       ELSIF (#tempEnable = FALSE) AND (#statEnableOld = TRUE) THEN // Disable FB 
           #statFBState := #FB_STATE_DISABLING;
       ELSIF (#statStatus = #STATUS_FIRST_CALL) THEN // Set status identifier of subsequent call
           #statStatus := #STATUS_SUBSEQUENT_CALL;
       END_IF;

       // Edge detection 'enable' input
       #statEnableOld := #tempEnable;
   END_REGION ENABLING/DISABLING

   IF (#statStatus = #STATUS_NO_CALL) THEN // Nothing to do -> End here to reduce "system load"
       RETURN;
   END_IF;

   REGION STATE_MACHINE_FUNCTION_BLOCK_TCP
       CASE #statFBState OF // State machine of FB
           #FB_STATE_NO_PROCESSING: // No processing active (Note: this state must always be present and left empty)
               ;

           #FB_STATE_VALIDATE_INPUT: // Enabling active
               REGION EVALUATE CONNECTION PARAMETERS
                   // Determine if host is domain name or IP address
                   #statConnParam.isQDN := NOT "IsIPAddress"(address := #connParam.broker, ipAddress => #statConnParam.paramIP.ConnPara.RemoteAddress);

                   IF #statConnParam.isQDN THEN // Broker address is a hostname
                       IF #connParam.broker[LEN(#connParam.broker)] = '.' THEN
                           #statConnParam.paramQDN.ConnPara.RemoteQDN := #connParam.broker;
                       ELSE
                           #statConnParam.paramQDN.ConnPara.RemoteQDN := CONCAT(IN1 := #connParam.broker, IN2 := '.');
                       END_IF;

                       #statConnParam.paramQDN.ConnPara.InterfaceId := #connParam.hwId;
                       #statConnParam.paramQDN.ConnPara.ID := #connParam.connId;
                       #statConnParam.paramQDN.ConnPara.ActiveEstablished := TRUE;
                       #statConnParam.paramQDN.ConnPara.RemotePort := #connParam."port";
                   ELSE // Broker address is an IP address
                       #statConnParam.paramIP.ConnPara.InterfaceId := #connParam.hwId;
                       #statConnParam.paramIP.ConnPara.ID := #statConnParam.paramQDN.ConnPara.ID := #connParam.connId;
                       #statConnParam.paramIP.ConnPara.ActiveEstablished := TRUE;
                       #statConnParam.paramIP.ConnPara.RemotePort := #connParam."port";
                   END_IF;

                   IF #connParam.tls.enableTls THEN
                       IF #statConnParam.isQDN THEN
                           #statConnParam.paramQDN.ActivateSecureConn := TRUE;
                           #statConnParam.paramQDN.ExtTLSCapabilities.%X0 := #connParam.tls.validateServerIdentity;
                           #statConnParam.paramQDN.TLSServerCertRef := #connParam.tls.brokerCert;
                           #statConnParam.paramQDN.TLSClientCertRef := #connParam.tls.clientCert;
                       ELSE
                           #statConnParam.paramIP.ActivateSecureConn := TRUE;
                           #statConnParam.paramIP.ExtTLSCapabilities.%X0 := #connParam.tls.validateServerIdentity;
                           #statConnParam.paramIP.TLSServerCertRef := #connParam.tls.brokerCert;
                           #statConnParam.paramIP.TLSClientCertRef := #connParam.tls.clientCert;
                       END_IF;
                   ELSE
                       IF #statConnParam.isQDN THEN
                           #statConnParam.paramQDN.ActivateSecureConn := FALSE;
                       ELSE
                           #statConnParam.paramIP.ActivateSecureConn := FALSE;
                       END_IF;
                   END_IF;
               END_REGION EVALUATE CONNECTION PARAMETERS

               REGION FB_VALIDATE_INPUT     
                   // Check Input variables:
                   #tempMaxWillMsgLen := ABS(UPPER_BOUND(ARR := #willMsgPayload, DIM := #ONE_DIMENSION) - LOWER_BOUND(ARR := #willMsgPayload, DIM := #ONE_DIMENSION)) + #ARRAY_LEN_OFFSET_PLUS_1;

                   // Check Client ID len Must be > 0 
                   IF LEN(#clientIdentifier) <= #LEN_NULL THEN
                       #statStatus := #ERR_CLIENT_ID_NULL; // Set correct status that identifies error clearly
                       #statSubfunctionStatus := #ERR_CLIENT_ID_NULL; // Status or return value of called FBs, FCs and system blocks
                       #statFBErrorState := #statFBState; // Set error state number for diagnostic 
                       #statErrorUserCleared := TRUE;

                       // Verify Will next
                   ELSIF #tempMaxWillMsgLen < #willMsgLen THEN
                       #statStatus := #ERR_CNT_EXCEEDS_ARRAY_DIMENSION; // Set correct status that identifies error clearly
                       #statSubfunctionStatus := #ERR_CNT_EXCEEDS_ARRAY_DIMENSION; // Status or return value of called FBs, FCs and system blocks
                       #statFBErrorState := #statFBState; // Set error state number for diagnostic 
                       #statErrorUserCleared := TRUE;

                       // Check Will QoS
                   ELSIF #qos > #MQTT_QOS_2 THEN
                       #statStatus := #ERR_QOS_INVALID; // Set correct status that identifies error clearly
                       #statSubfunctionStatus := #ERR_QOS_INVALID; // Status or return value of called FBs, FCs and system blocks
                       #statFBErrorState := #statFBState; // Set error state number for diagnostic 
                       #statErrorUserCleared := TRUE;

                       // Check KeepAlive
                   ELSIF (#connParam.keepAlive < #THREE_SECONDS) // IF Set to 1 or 2 seconds..
                       AND (#connParam.keepAlive > 0)
                   THEN
                       #statStatus := #ERR_KEEPALIVE_INVALID; // Set correct status that identifies error clearly
                       #statSubfunctionStatus := #ERR_KEEPALIVE_INVALID; // Status or return value of called FBs, FCs and system blocks
                       #statFBErrorState := #statFBState; // Set error state number for diagnostic 
                       #statErrorUserCleared := TRUE;

                   ELSE
                       // Set Params for connection
                       // Set Client Id
                       #statWillQos := #qos;
                       // Set Retain
                       #statWillRetain := #retain;
                       // Will message cnt
                       #statWillMessageCnt := #willMsgLen;

                       // Keepalive
                       IF #connParam.keepAlive = 0 THEN
                           #statMqttKeepAliveUsed := FALSE;
                       ELSE
                           #statMqttKeepAliveUsed := TRUE;
                           // KeepAliveTImer is set to ((Keep Alive converted to seconds) - 2s)
                           #statMqttKeepAliveTime := UINT_TO_TIME((#connParam.keepAlive * #UINT_CONST_1000 - #TWO_SECONDS));
                       END_IF;

                       // rdy to enable TCON
                       #statTsendcEnable := TRUE;
                       #statEnableTimerCommandWatchdog := TRUE;
                       #statFBState := #FB_STATE_TCP_CONNECTING;
                   END_IF;
               END_REGION FB_VALIDATE_INPUT

           #FB_STATE_TCP_CONNECTING: // Wait for TCP to be established
               REGION FB_TCP_CONNECTING
                   // Check process:
                   IF #tempTsendcError = TRUE THEN // when error:
                       #statTsendcEnable := FALSE; // disable TsendC
                       #statEnableTimerCommandWatchdog := FALSE;
                       #statStatus := #ERR_TCON_FAILED; // Set correct status that identifies error clearly
                       #statSubfunctionStatus := #tempTsendcStatus; // Status or return value of called FBs, FCs and system blocks
                       #statFBErrorState := #statFBState; // Set error state number for diagnostic 
                       #statErrorUserCleared := TRUE;

                   ELSIF #tempTsendcStatus = #TSENDC_EST_OK THEN // when successfull:
                       // Communication connection established.
                       #statEnableTimerCommandWatchdog := FALSE;
                       // Monitor Connection
                       #statFBState := #FB_STATE_OPERATING_MONITOR_TCP;
                       // Begin MQTT Connection
                       #statMqttConnectState := #MQTT_CONNECT_STATE_BUILD_PACKET;
                       // set status
                       #statStatus := #STATUS_MQTT_CONNECTING;

                   ELSIF #instTimerCommandWatchdog.Q THEN
                       #statTsendcEnable := FALSE; // disable TsendC
                       #statEnableTimerCommandWatchdog := FALSE;
                       #statStatus := #ERR_TCON_TIMEOUT; // Set correct status that identifies error clearly
                       #statSubfunctionStatus := #ERR_TCON_TIMEOUT; // Status or return value of called FBs, FCs and system blocks
                       #statFBErrorState := #statFBState; // Set error state number for diagnostic 
                       #statErrorUserCleared := TRUE;
                   END_IF;
               END_REGION FB_TCP_CONNECTING

           #FB_STATE_OPERATING_MONITOR_TCP: // Processing active
               REGION FB_OPERATING_MONITOR_TCP
                   // Reset Status on Msg Output - will be set when a new message is completly processed and ready at outputs.
                   #statRcvMsgStatus := #MSG_DECODE_STATUS_NO_NEW_MSG;
                   // Reset TsendC Req from last  cycle Request:
                   #statTsendcReq := FALSE;

                   // Monitor Connection - if disconnect occured:
                   IF ((#tempTsendcStatus > #TSENDC_COM_CLOSED AND #tempTsendcStatus < #TSENDC_EST_OK) // Status connection interupt
                       OR #tempTsendcError = TRUE) // Or error
                       AND #tempTrcvNdr = FALSE // And no new data (to see if broker send information why connection was interrupted)
                   THEN
                       REGION CONNECTION_INTERRUPTED
                           // Status reconnecting
                           // SET MQTT to no operation
                           #statMqttConnectState := #MQTT_CONNECT_STATE_NO_PROCESSING;
                           #statMqttCommandState := #MQTT_COMMAND_STATE_NO_PROCESSING;
                           #statRcvMsgDecodeState := #MSG_DECODE_STATE_NO_PROCESSING;
                           // Reset PUBACK / PUBREC / PUBCOMP
                           #statSendPubAckMsg :=
                           #statSendPubRecMsg :=
                           #statSendPubCompMsg := FALSE;
                           // reset Done bit if still set, regardless of input:
                           #statDone := FALSE;
                           // reset Watchdog
                           #statEnableTimerCommandWatchdog := FALSE;
                           // reset headerEncode
                           #statPacketHeaderEncodeDone := FALSE;
                           // set error  information
                           #statStatus := #ERR_TCP_RECONNECTING; // Set correct status that identifies error clearly
                           #statSubfunctionStatus := #tempTsendcStatus;// Status or return value of called FBs, FCs and system blocks
                           #statFBErrorState := #statFBState; // Set error state number for diagnostic 
                           #statErrorAutoCleared := TRUE;
                           // Wait for reconect - next state
                           #statFBState := #FB_STATE_TCP_RECONNECTING;
                       END_REGION REGION CONNECTION_INTERRUPTED
                   ELSE
                       // Connection is OK
                       // Sending and receiving works 
                       // Check Trcv Buffer for new Data
                       IF #tempTrcvNdr THEN
                           REGION TRCV_NEW_DATA
                               // Evaluate the TrcvBuffer, reset buffer pos to start
                               #tempTrcvBufferPos := 0;

                               // Parse the whole RCV Buffer
                               // While there is data to be processed
                               WHILE ((#tempTrcvBufferPos = UDINT_TO_DINT(#tempTrcvRcvdLen) AND #statRcvMsgDecodeState = #MSG_DECODE_STATE_COMPLETED)
                                   OR #tempTrcvBufferPos < UDINT_TO_DINT(#tempTrcvRcvdLen))
                               DO
                                   // Parse the whole RCV Buffer, check wether header or decoding
                                   IF #statRcvMsgDecodeState = #MSG_DECODE_STATE_NO_PROCESSING THEN
                                       // If no decoding is in progress, look for new message header
                                       #tempRcvMsgTypeCase := #statRcvBuffer[#tempTrcvBufferPos] AND #BIT_MASK_HIGHBITS;
                                   ELSE
                                       // Decode is in progress, go directly to decoding
                                       #tempRcvMsgTypeCase := #MQTT_MSG_DECODING;
                                   END_IF;

                                   CASE #tempRcvMsgTypeCase OF

                                       #MQTT_MSG_TYPE_CONNACK:
                                           REGION RECEIVED_CONACK_PACKET
                                               // Check all CONNACK packet is inside the receive buffer
                                               IF #tempTrcvBufferPos + #BYTE_SIZE_CONNACK <= #MAX_BUFFER_LEN_RCV THEN
                                                   #tempTrcvBufferPos += 1;
                                                   IF #statRcvBuffer[#tempTrcvBufferPos] = #REMAINING_LEN_2 THEN // remainng Length must be 2;
                                                       #tempTrcvBufferPos += 1;
                                                       // byte one is 0000 000X where X is if Session was set, so depending on clean session or not evaluate answer of server
                                                       #statSessionPresent := #statRcvBuffer[#tempTrcvBufferPos] <> #MQTT_NO_SESSION_PRESENT;
                                                       IF (#cleanSession AND NOT #statSessionPresent)
                                                           OR NOT #cleanSession
                                                       THEN
                                                           #tempTrcvBufferPos += 1;
                                                           // VALID Answer, check code
                                                           IF #statRcvBuffer[#tempTrcvBufferPos] = #MQTT_CONNACK_ACCEPTED THEN
                                                               // All good
                                                               #tempTrcvBufferPos += 1;
                                                               #tempMqttConnAckRcvStatus := #RESPONSE_GOOD; // evaluate in MQTT StateMachine Below the response
                                                           ELSE
                                                               // NOT VALID CONNACK from server shows session has a bad return code
                                                               #statStatus := #ERR_MQTT_CONNACK_RETURN_CODE_INVALID; // Set correct status that identifies error clearly
                                                               #statSubfunctionStatus := #statRcvBuffer[#tempTrcvBufferPos]; // Status or return value of called FBs, FCs and system blocks
                                                               #statFBErrorState := #statFBState; // Set error state number for diagnostic 
                                                               #statErrorUserCleared := TRUE;
                                                               // Exit loop
                                                               EXIT;
                                                           END_IF;
                                                       ELSE
                                                           // NOT VALID, CONNACK from server shows session present
                                                           #statStatus := #ERR_MQTT_CONNACK_INVALID_SESSION_FLAG; // Set correct status that identifies error clearly
                                                           #statSubfunctionStatus := #ERR_MQTT_CONNACK_INVALID_SESSION_FLAG; // Status or return value of called FBs, FCs and system blocks
                                                           #statFBErrorState := #statFBState; // Set error state number for diagnostic 
                                                           #statErrorUserCleared := TRUE;
                                                           // Exit loop
                                                           EXIT;
                                                       END_IF;
                                                   ELSE // We got a CONNACK packet, but remaining length was not 2 (Error)
                                                       #statStatus := #ERR_MQTT_REM_LEN_INVALID; // Set correct status that identifies error clearly
                                                       #statSubfunctionStatus := #ERR_MQTT_REM_LEN_INVALID; // Status or return value of called FBs, FCs and system blocks
                                                       #statFBErrorState := #statFBState; // Set error state number for diagnostic 
                                                       #statErrorUserCleared := TRUE;
                                                       // Exit loop
                                                       EXIT;
                                                   END_IF;
                                               ELSE
                                                   // If the CONNACK packed is not fully inside the receive buffer, finish processing
                                                   #statStatus := #ERR_MSG_SKIPPED; // Set correct status that identifies error clearly
                                                   #statSubfunctionStatus := #ERR_MSG_SKIPPED; // Status or return value of called FBs, FCs and system blocks
                                                   #statFBErrorState := #statFBState; // Set error state number for diagnostic 
                                                   #statErrorUserCleared := TRUE;
                                                   // Exit loop
                                                   EXIT;
                                               END_IF;
                                           END_REGION RECEIVED_CONACK_PACKET

                                       #MQTT_MSG_TYPE_PINGRESP:
                                           REGION RECEIVED_PINGRESP_PACKET
                                               // Check all PINGRESP packet is inside the receive buffer
                                               IF #tempTrcvBufferPos + #BYTE_SIZE_PINGRESP <= #MAX_BUFFER_LEN_RCV THEN
                                                   #tempTrcvBufferPos += 1;
                                                   IF #statRcvBuffer[#tempTrcvBufferPos] = #REMAINING_LEN_0 THEN // remainng Length must be 0;
                                                       #tempTrcvBufferPos += 1;
                                                       #tempMqttPingRspRcv := #RESPONSE_GOOD; // evaluate in MQTT StateMachine Below the response
                                                   ELSE // We got a Pingrsp packet, but remaining length was not 0 (Error)
                                                       #statStatus := #ERR_MQTT_REM_LEN_INVALID; // Set correct status that identifies error clearly
                                                       #statSubfunctionStatus := #ERR_MQTT_REM_LEN_INVALID; // Status or return value of called FBs, FCs and system blocks
                                                       #statFBErrorState := #statFBState; // Set error state number for diagnostic 
                                                       #statErrorAutoCleared := TRUE;
                                                       // Exit loop
                                                       EXIT;
                                                   END_IF;
                                               ELSE
                                                   // If the PINGRESP packed is not fully inside the receive buffer, finish processing
                                                   #statStatus := #ERR_MSG_SKIPPED; // Set correct status that identifies error clearly
                                                   #statSubfunctionStatus := #ERR_MSG_SKIPPED; // Status or return value of called FBs, FCs and system blocks
                                                   #statFBErrorState := #statFBState; // Set error state number for diagnostic 
                                                   #statErrorAutoCleared := TRUE;
                                                   // Exit loop
                                                   EXIT;
                                               END_IF;
                                           END_REGION RECEIVED_PINGRESP_PACKET

                                       #MQTT_MSG_TYPE_PUBACK:
                                           REGION RECEIVED_PUBACK_PACKET
                                               // Check all PUBACK packet is inside the receive buffer
                                               IF #tempTrcvBufferPos + #BYTE_SIZE_PUBACK <= #MAX_BUFFER_LEN_RCV THEN
                                                   #tempTrcvBufferPos += 1;
                                                   IF #statRcvBuffer[#tempTrcvBufferPos] = #REMAINING_LEN_2 THEN// remaining Length must be 2;
                                                       #tempTrcvBufferPos += 1;
                                                       #tempWordForSliceAddress := UINT_TO_WORD(#statPacketId);
                                                       IF #statRcvBuffer[#tempTrcvBufferPos] = #tempWordForSliceAddress.%B1 THEN
                                                           #tempTrcvBufferPos += 1;
                                                           IF #statRcvBuffer[#tempTrcvBufferPos] = #tempWordForSliceAddress.%B0 THEN
                                                               #tempTrcvBufferPos += 1;
                                                               #tempMqttPubAckRcv := #RESPONSE_GOOD;
                                                           ELSE
                                                               #tempTrcvBufferPos += 1;
                                                               #tempMqttPubAckRcv := #RESPONSE_PACKET_ID_INVALID;
                                                           END_IF;
                                                       ELSE
                                                           #tempTrcvBufferPos += 1;
                                                           #tempMqttPubAckRcv := #RESPONSE_PACKET_ID_INVALID;
                                                       END_IF;
                                                   ELSE
                                                       #statStatus := #ERR_MQTT_REM_LEN_INVALID; // Set correct status that identifies error clearly
                                                       #statSubfunctionStatus := #ERR_MQTT_REM_LEN_INVALID; // Status or return value of called FBs, FCs and system blocks
                                                       #statFBErrorState := #statFBState; // Set error state number for diagnostic 
                                                       #statErrorAutoCleared := TRUE;
                                                       // Exit loop
                                                       EXIT;
                                                   END_IF;
                                               ELSE
                                                   // If the PUBACK packed is not fully inside the receive buffer, finish processing
                                                   #statStatus := #ERR_MSG_SKIPPED; // Set correct status that identifies error clearly
                                                   #statSubfunctionStatus := #ERR_MSG_SKIPPED; // Status or return value of called FBs, FCs and system blocks
                                                   #statFBErrorState := #statFBState; // Set error state number for diagnostic 
                                                   #statErrorAutoCleared := TRUE;
                                                   // Exit loop
                                                   EXIT;
                                               END_IF;
                                           END_REGION RECEIVED_PUBACK_PACKET

                                       #MQTT_MSG_TYPE_PUBREC:
                                           REGION RECEIVED_PUBREC_PACKET
                                               // Check all PUBREC packet is inside the receive buffer
                                               IF #tempTrcvBufferPos + #BYTE_SIZE_PUBREC <= #MAX_BUFFER_LEN_RCV THEN
                                                   #tempTrcvBufferPos += 1;
                                                   IF #statRcvBuffer[#tempTrcvBufferPos] = #REMAINING_LEN_2 THEN// remainng Length must be 2;
                                                       #tempTrcvBufferPos += 1;
                                                       #tempWordForSliceAddress := UINT_TO_WORD(#statPacketId);
                                                       IF #statRcvBuffer[#tempTrcvBufferPos] = #tempWordForSliceAddress.%B1 THEN
                                                           #tempTrcvBufferPos += 1;
                                                           IF #statRcvBuffer[#tempTrcvBufferPos] = #tempWordForSliceAddress.%B0 THEN
                                                               #tempTrcvBufferPos += 1;
                                                               #statMqttPubRecRcv := #RESPONSE_GOOD;
                                                           ELSE
                                                               #tempTrcvBufferPos += 1;
                                                               #statMqttPubRecRcv := #RESPONSE_PACKET_ID_INVALID;
                                                           END_IF;
                                                       ELSE
                                                           #tempTrcvBufferPos += 1;
                                                           #statMqttPubRecRcv := #RESPONSE_PACKET_ID_INVALID;
                                                       END_IF;
                                                   ELSE
                                                       #statStatus := #ERR_MQTT_REM_LEN_INVALID; // Set correct status that identifies error clearly
                                                       #statSubfunctionStatus := #ERR_MQTT_REM_LEN_INVALID; // Status or return value of called FBs, FCs and system blocks
                                                       #statFBErrorState := #statFBState; // Set error state number for diagnostic 
                                                       #statErrorAutoCleared := TRUE;
                                                       // Exit loop
                                                       EXIT;
                                                   END_IF;
                                               ELSE
                                                   // If the PUBREC packed is not fully inside the receive buffer, finish processing
                                                   #statStatus := #ERR_MSG_SKIPPED; // Set correct status that identifies error clearly
                                                   #statSubfunctionStatus := #ERR_MSG_SKIPPED; // Status or return value of called FBs, FCs and system blocks
                                                   #statFBErrorState := #statFBState; // Set error state number for diagnostic 
                                                   #statErrorAutoCleared := TRUE;
                                                   // Exit loop
                                                   EXIT;
                                               END_IF;
                                           END_REGION RECEIVED_PUBREC_PACKET

                                       #MQTT_MSG_TYPE_PUBREL:
                                           REGION RECEIVED_PUBREL_PACKET
                                               // Check all PUBREL packet is inside the receive buffer
                                               IF #tempTrcvBufferPos + #BYTE_SIZE_PUBREL <= #MAX_BUFFER_LEN_RCV THEN
                                                   #tempTrcvBufferPos += 1;
                                                   IF #statRcvBuffer[#tempTrcvBufferPos] = #REMAINING_LEN_2 THEN // Remaining Length must be 2
                                                       #tempTrcvBufferPos += 1;
                                                       #tempWordForSliceAddress.%B1 := #statRcvBuffer[#tempTrcvBufferPos];
                                                       #tempTrcvBufferPos += 1;
                                                       #tempWordForSliceAddress.%B0 := #statRcvBuffer[#tempTrcvBufferPos];
                                                       #tempTrcvBufferPos += 1;
                                                       #statRelPacketId := #EMPTY_WORD;

                                                       // Is there a QoS2 subscribed message to be released
                                                       FOR #tempStorageIndex := 0 TO #MAX_BUFFER_LEN_QOS2 DO
                                                           IF #statRcvPacketIdStorage[#tempStorageIndex] = #tempWordForSliceAddress THEN
                                                               #statRelPacketId := #statRcvPacketIdStorage[#tempStorageIndex];
                                                               EXIT;
                                                           END_IF;
                                                       END_FOR;

                                                       IF #statRelPacketId <> #EMPTY_WORD THEN
                                                           #statMqttPubRelRcv := #RESPONSE_GOOD;

                                                           // Get maximum payload size
                                                           #tempReceivedMsgDataArrayTotalLen := ABS(UPPER_BOUND(ARR := #receivedMsgPayload, DIM := #ONE_DIMENSION) - LOWER_BOUND(ARR := #receivedMsgPayload, DIM := #ONE_DIMENSION)) + #ARRAY_LEN_OFFSET_PLUS_1;
                                                           IF #tempReceivedMsgDataArrayTotalLen <= #MAX_BUFFER_LEN_RCV + #ARRAY_LEN_OFFSET_PLUS_1 THEN
                                                               // The limit is given by the payload output array
                                                               IF #statRcvMsgPayloadLenStorage[#tempStorageIndex] > #tempReceivedMsgDataArrayTotalLen THEN
                                                                   #statRcvMsgDataLen := DINT_TO_UDINT(#tempReceivedMsgDataArrayTotalLen);
                                                               ELSE
                                                                   #statRcvMsgDataLen := #statRcvMsgPayloadLenStorage[#tempStorageIndex];
                                                               END_IF;
                                                           ELSE
                                                               // The limit is given by the QoS2 buffer array
                                                               IF #statRcvMsgPayloadLenStorage[#tempStorageIndex] > #MAX_BUFFER_LEN_RCV + #ARRAY_LEN_OFFSET_PLUS_1 THEN
                                                                   #statRcvMsgDataLen := #MAX_BUFFER_LEN_RCV + #ARRAY_LEN_OFFSET_PLUS_1;
                                                               ELSE
                                                                   #statRcvMsgDataLen := #statRcvMsgPayloadLenStorage[#tempStorageIndex];
                                                               END_IF;
                                                           END_IF;

                                                           MOVE_BLK(IN := #statRcvPayloadStorage[#tempStorageIndex, 0],
                                                                    COUNT := #statRcvMsgDataLen,
                                                                    OUT => #receivedMsgPayload[LOWER_BOUND(ARR := #receivedMsgPayload, DIM := #ONE_DIMENSION)]);

                                                           #receivedTopic := #statRcvTopicStorage[#tempStorageIndex]; // Send Payload to in/out 
                                                           #statRcvPacketIdStorage[#tempStorageIndex] := #EMPTY_WORD; // release stored PacketId
                                                           IF #statRcvMsgDataLen < #statRcvMsgPayloadLenStorage[#tempStorageIndex] THEN
                                                               #statRcvMsgInternalStatus := #MSG_DECODE_STATUS_PAYLOAD_TOO_LONG;
                                                           ELSE
                                                               #statRcvMsgInternalStatus := #MSG_DECODE_STATUS_NEW_MSG_OK;
                                                           END_IF;
                                                           #statSendPubCompMsg := TRUE;
                                                       ELSE
                                                           #tempTrcvBufferPos += 1;
                                                           #statMqttPubRelRcv := #RESPONSE_PACKET_ID_INVALID;
                                                       END_IF;
                                                   ELSE
                                                       #statStatus := #ERR_MQTT_REM_LEN_INVALID; // Set correct status that identifies error clearly
                                                       #statSubfunctionStatus := #ERR_MQTT_REM_LEN_INVALID; // Status or return value of called FBs, FCs and system blocks
                                                       #statFBErrorState := #statFBState; // Set error state number for diagnostic 
                                                       #statErrorAutoCleared := TRUE;
                                                       // Exit loop
                                                       EXIT;
                                                   END_IF;
                                               ELSE
                                                   // If the PUBREL packed is not fully inside the receive buffer, finish processing
                                                   #statStatus := #ERR_MSG_SKIPPED; // Set correct status that identifies error clearly
                                                   #statSubfunctionStatus := #ERR_MSG_SKIPPED; // Status or return value of called FBs, FCs and system blocks
                                                   #statFBErrorState := #statFBState; // Set error state number for diagnostic 
                                                   #statErrorAutoCleared := TRUE;
                                                   // Exit loop
                                                   EXIT;
                                               END_IF;
                                           END_REGION RECEIVED_PUBREL_PACKET      

                                       #MQTT_MSG_TYPE_PUBCOMP:
                                           REGION RECEIVED_PUBCOMP_PACKET
                                               // Check all PUBCOMP packet is inside the receive buffer
                                               IF #tempTrcvBufferPos + #BYTE_SIZE_PUBCOMP <= #MAX_BUFFER_LEN_RCV THEN
                                                   #tempTrcvBufferPos += 1;
                                                   IF #statRcvBuffer[#tempTrcvBufferPos] = #REMAINING_LEN_2 THEN // remaining Length must be 2
                                                       #tempTrcvBufferPos += 1;
                                                       #tempWordForSliceAddress := UINT_TO_WORD(#statPacketId);
                                                       IF #statRcvBuffer[#tempTrcvBufferPos] = #tempWordForSliceAddress.%B1 THEN
                                                           #tempTrcvBufferPos += 1;
                                                           IF #statRcvBuffer[#tempTrcvBufferPos] = #tempWordForSliceAddress.%B0 THEN
                                                               #tempTrcvBufferPos += 1;
                                                               #tempMqttPubCompRcv := #RESPONSE_GOOD;
                                                           ELSE
                                                               #tempTrcvBufferPos += 1;
                                                               #tempMqttPubCompRcv := #RESPONSE_PACKET_ID_INVALID;
                                                           END_IF;
                                                       ELSE
                                                           #tempTrcvBufferPos += 1;
                                                           #tempMqttPubCompRcv := #RESPONSE_PACKET_ID_INVALID;
                                                       END_IF;
                                                   ELSE
                                                       #statStatus := #ERR_MQTT_REM_LEN_INVALID; // Set correct status that identifies error clearly
                                                       #statSubfunctionStatus := #ERR_MQTT_REM_LEN_INVALID; // Status or return value of called FBs, FCs and system blocks
                                                       #statFBErrorState := #statFBState; // Set error state number for diagnostic 
                                                       #statErrorAutoCleared := TRUE;
                                                       // Exit loop
                                                       EXIT;
                                                   END_IF;
                                               ELSE
                                                   // If the PUBCOMP packed is not fully inside the receive buffer, finish processing
                                                   #statStatus := #ERR_MSG_SKIPPED; // Set correct status that identifies error clearly
                                                   #statSubfunctionStatus := #ERR_MSG_SKIPPED; // Status or return value of called FBs, FCs and system blocks
                                                   #statFBErrorState := #statFBState; // Set error state number for diagnostic 
                                                   #statErrorAutoCleared := TRUE;
                                                   // Exit loop
                                                   EXIT;
                                               END_IF;
                                           END_REGION RECEIVED_PUBCOMP_PACKET

                                       #MQTT_MSG_TYPE_SUBACK:
                                           REGION RECEIVED_SUBACK_PACKET
                                               // Check all SUBACK packet is inside the receive buffer
                                               IF #tempTrcvBufferPos + #BYTE_SIZE_SUBACK <= #MAX_BUFFER_LEN_RCV THEN
                                                   #tempTrcvBufferPos += 1;
                                                   IF #statRcvBuffer[#tempTrcvBufferPos] = #REMAINING_LEN_3 THEN // remaining Length must be 3
                                                       #tempTrcvBufferPos += 1;
                                                       #tempWordForSliceAddress := UINT_TO_WORD(#statPacketId);
                                                       IF #statRcvBuffer[#tempTrcvBufferPos] = #tempWordForSliceAddress.%B1 THEN
                                                           #tempTrcvBufferPos += 1;
                                                           IF #statRcvBuffer[#tempTrcvBufferPos] = #tempWordForSliceAddress.%B0 THEN
                                                               #tempTrcvBufferPos += 1;
                                                               IF #statRcvBuffer[#tempTrcvBufferPos] = #SUBSCRIBE_FAILURE THEN
                                                                   #tempTrcvBufferPos += 1;
                                                                   #tempMqttSubAckRcv := #RESPONSE_SUBSCRIBE_FAILED;
                                                               ELSE
                                                                   #tempTrcvBufferPos += 1;
                                                                   #tempMqttSubAckRcv := #RESPONSE_GOOD;
                                                               END_IF;
                                                           ELSE
                                                               #tempTrcvBufferPos += 1;
                                                               #tempMqttSubAckRcv := #RESPONSE_PACKET_ID_INVALID;
                                                           END_IF;
                                                       ELSE
                                                           #tempTrcvBufferPos += 1;
                                                           #tempMqttSubAckRcv := #RESPONSE_PACKET_ID_INVALID;
                                                       END_IF;
                                                   ELSE
                                                       #statStatus := #ERR_MQTT_REM_LEN_INVALID; // Set correct status that identifies error clearly
                                                       #statSubfunctionStatus := #ERR_MQTT_REM_LEN_INVALID; // Status or return value of called FBs, FCs and system blocks
                                                       #statFBErrorState := #statFBState; // Set error state number for diagnostic 
                                                       #statErrorAutoCleared := TRUE;
                                                       // Exit loop
                                                       EXIT;
                                                   END_IF;
                                               ELSE
                                                   // If the SUBACK packed is not fully inside the receive buffer, finish processing
                                                   #statStatus := #ERR_MSG_SKIPPED; // Set correct status that identifies error clearly
                                                   #statSubfunctionStatus := #ERR_MSG_SKIPPED; // Status or return value of called FBs, FCs and system blocks
                                                   #statFBErrorState := #statFBState; // Set error state number for diagnostic 
                                                   #statErrorAutoCleared := TRUE;
                                                   // Exit loop
                                                   EXIT;
                                               END_IF;
                                           END_REGION RECEIVED_SUBACK_PACKET

                                       #MQTT_MSG_TYPE_UNSUBACK:
                                           REGION RECEIVED_UNSUBACK_PACKET
                                               // Check all UNSUBACK packet is inside the receive buffer
                                               IF #tempTrcvBufferPos + #BYTE_SIZE_UNSUBACK <= #MAX_BUFFER_LEN_RCV THEN
                                                   #tempTrcvBufferPos += 1;
                                                   IF #statRcvBuffer[#tempTrcvBufferPos] = #REMAINING_LEN_2 THEN // remaining Length must be 2
                                                       #tempTrcvBufferPos += 1;
                                                       #tempWordForSliceAddress := UINT_TO_WORD(#statPacketId);
                                                       IF #statRcvBuffer[#tempTrcvBufferPos] = #tempWordForSliceAddress.%B1 THEN
                                                           #tempTrcvBufferPos += 1;
                                                           IF #statRcvBuffer[#tempTrcvBufferPos] = #tempWordForSliceAddress.%B0 THEN
                                                               #tempTrcvBufferPos += 1;
                                                               #tempMqttUnSubAckRcv := #RESPONSE_GOOD;
                                                           ELSE
                                                               #tempTrcvBufferPos += 1;
                                                               #tempMqttUnSubAckRcv := #RESPONSE_PACKET_ID_INVALID;
                                                           END_IF;
                                                       ELSE
                                                           #tempTrcvBufferPos += 1;
                                                           #tempMqttUnSubAckRcv := #RESPONSE_PACKET_ID_INVALID;
                                                       END_IF;
                                                   ELSE
                                                       #statStatus := #ERR_MQTT_REM_LEN_INVALID; // Set correct status that identifies error clearly
                                                       #statSubfunctionStatus := #ERR_MQTT_REM_LEN_INVALID; // Status or return value of called FBs, FCs and system blocks
                                                       #statFBErrorState := #statFBState; // Set error state number for diagnostic 
                                                       #statErrorAutoCleared := TRUE;
                                                       // Exit loop
                                                       EXIT;
                                                   END_IF;
                                               ELSE
                                                   // If the UNSUBACK packed is not fully inside the receive buffer, finish processing
                                                   #statStatus := #ERR_MSG_SKIPPED; // Set correct status that identifies error clearly
                                                   #statSubfunctionStatus := #ERR_MSG_SKIPPED; // Status or return value of called FBs, FCs and system blocks
                                                   #statFBErrorState := #statFBState; // Set error state number for diagnostic 
                                                   #statErrorAutoCleared := TRUE;
                                                   // Exit loop
                                                   EXIT;
                                               END_IF;
                                           END_REGION RECEIVED_UNSUBACK_PACKET

                                       #MQTT_MSG_TYPE_PUBLISH:
                                           REGION RECEIVED_PUBLISH_PACKET
                                               // Received a message, start process.
                                               #tempMultiplierToDecode := #INIT_UDINT_1;
                                               #statRcvMsgTotalLen := 0;
                                               #statRcvMsgTopicLen := 0;
                                               #statRcvMsgPayloadLen := 0;

                                               // Check that at least the reamaining length and topic size of the PUBLISH packet is inside the receive buffer
                                               IF #tempTrcvBufferPos + #BYTE_SIZE_PUBLISH <= #MAX_BUFFER_LEN_RCV THEN
                                                   // Check and store QoS for later use
                                                   IF (#statRcvBuffer[#tempTrcvBufferPos] AND #BIT_MASK_QOS) = #MQTT_MSG_QOS0 THEN
                                                       #statRcvMsgQoS := #MQTT_QOS_0;
                                                   ELSIF (#statRcvBuffer[#tempTrcvBufferPos] AND #BIT_MASK_QOS) = #MQTT_MSG_QOS1 THEN
                                                       #statRcvMsgQoS := #MQTT_QOS_1;
                                                   ELSIF (#statRcvBuffer[#tempTrcvBufferPos] AND #BIT_MASK_QOS) = #MQTT_MSG_QOS2 THEN
                                                       #statRcvMsgQoS := #MQTT_QOS_2;
                                                   ELSIF (#statRcvBuffer[#tempTrcvBufferPos] AND #BIT_MASK_QOS) = #MQTT_MSG_QOS_BAD THEN
                                                       #statStatus := #ERR_MQTT_MALFORMED_QOS_RECEIVED; // Set correct status that identifies error clearly
                                                       #statSubfunctionStatus := #ERR_MQTT_MALFORMED_QOS_RECEIVED; // Status or return value of called FBs, FCs and system blocks
                                                       #statFBErrorState := #statFBState; // Set error state number for diagnostic 
                                                       #statErrorAutoCleared := TRUE;
                                                       // Exit loop
                                                       EXIT;
                                                   END_IF;

                                                   // Calculate total publish len (topic,packetid,payload)
                                                   REPEAT
                                                       #tempTrcvBufferPos += 1; // Increment
                                                       #statRcvMsgTotalLen += BYTE_TO_UDINT((#statRcvBuffer[#tempTrcvBufferPos] AND #DEFAULT_MULTIPLIER_BYTE_127)) * #tempMultiplierToDecode;
                                                       #tempMultiplierToDecode *= #SEND_LEN_MULTIPLIER_UDINT_128;
                                                       IF #tempMultiplierToDecode > #MAX_ALLOWED_PACKET_SIZE THEN
                                                           // Throw error here // Malformed remain length.
                                                           #statStatus := #ERR_MQTT_REM_LEN_INVALID; // Set correct status that identifies error clearly
                                                           #statSubfunctionStatus := #ERR_MQTT_REM_LEN_INVALID; // Status or return value of called FBs, FCs and system blocks
                                                           #statFBErrorState := #statFBState; // Set error state number for diagnostic 
                                                           #statErrorAutoCleared := TRUE;
                                                           // Exit loop
                                                           EXIT;
                                                       END_IF;
                                                   UNTIL ((#statRcvBuffer[#tempTrcvBufferPos] AND UDINT_TO_BYTE(#SEND_LEN_MULTIPLIER_UDINT_128)) = 0)
                                                   END_REPEAT;

                                                   #tempTrcvBufferPos += 1; // Increment
                                                   // Save Topic Len
                                                   #tempWordForSliceAddress.%B1 := #statRcvBuffer[#tempTrcvBufferPos]; // MSB
                                                   #tempTrcvBufferPos += 1; // Increment
                                                   #tempWordForSliceAddress.%B0 := #statRcvBuffer[#tempTrcvBufferPos]; // LSB
                                                   #tempTrcvBufferPos += 1; // Increment
                                                   #statRcvMsgTopicLen := WORD_TO_UINT(#tempWordForSliceAddress);
                                                   // Set Payload len
                                                   IF #statRcvMsgQoS = #MQTT_QOS_0 THEN
                                                       // Payload Len is total Len minus topic len minus topic len info 
                                                       #statRcvMsgPayloadLen :=
                                                       #statDecodedPayloadLenght := #statRcvMsgTotalLen - #statRcvMsgTopicLen - #TWO_BYTE_LEN_INFO;
                                                   ELSE
                                                       // PayloadLen is total Len minus topic len minus topic len info minus packet Id len
                                                       #statRcvMsgPayloadLen :=
                                                       #statDecodedPayloadLenght := #statRcvMsgTotalLen - #statRcvMsgTopicLen - #TWO_BYTE_LEN_INFO - #TWO_BYTE_LEN_INFO;
                                                   END_IF;

                                                   // Select empty storage place if received publish message is received with QoS2
                                                   IF #statRcvMsgQoS = #MQTT_QOS_2 THEN
                                                       #statStoragePos := -1;
                                                       REPEAT
                                                           #statStoragePos += 1;
                                                           IF #statRcvPacketIdStorage[#statStoragePos] = #EMPTY_WORD THEN
                                                               EXIT;
                                                           END_IF;
                                                       UNTIL #statStoragePos = #MAX_BUFFER_LEN_QOS2
                                                       END_REPEAT;
                                                       IF #statStoragePos = -1 THEN
                                                           #statStatus := #ERR_CNT_QOS2_STORAGE_FULL; // Set correct status that identifies error clearly
                                                           #statSubfunctionStatus := #ERR_CNT_EXCEEDS_ARRAY_DIMENSION; // Status or return value of called FBs, FCs and system blocks
                                                           #statFBErrorState := #statFBState; // Set error state number for diagnostic 
                                                           #statErrorUserCleared := TRUE;
                                                           // Exit loop
                                                           EXIT;
                                                       END_IF;
                                                   END_IF;

                                                   // Clear Output message:
                                                   #receivedTopic := #EMPTY_WSTRING;
                                                   // Start Topic at first character
                                                   #statRcvMsgTopicPos := #FIRST_CHARACTER;
                                                   // Start RcvMsg at first array element
                                                   IF #statRcvMsgQoS = #MQTT_QOS_2 THEN
                                                       #statRcvMsgPayloadPos := 0;
                                                   ELSE
                                                       #statRcvMsgPayloadPos := LOWER_BOUND(ARR := #receivedMsgPayload, DIM := #ONE_DIMENSION);
                                                   END_IF;

                                                   // Start receiving with topic
                                                   #statRcvMsgDecodeState := #MSG_DECODE_STATE_TOPIC;

                                               ELSE
                                                   #statStatus := #ERR_MSG_SKIPPED; // Set correct status that identifies error clearly
                                                   #statSubfunctionStatus := #ERR_MSG_SKIPPED; // Status or return value of called FBs, FCs and system blocks
                                                   #statFBErrorState := #statFBState; // Set error state number for diagnostic 
                                                   #statErrorAutoCleared := TRUE;
                                                   // Exit loop
                                                   EXIT;
                                               END_IF;
                                           END_REGION RECEIVED_PUBLISH_PACKET

                                       #MQTT_MSG_DECODING:
                                           REGION RECEIVED_PACKET_DECODE

                                               CASE #statRcvMsgDecodeState OF
                                                   #MSG_DECODE_STATE_NO_PROCESSING: // No processing
                                                       ;

                                                   #MSG_DECODE_STATE_TOPIC:
                                                       // Decode topic
                                                       IF #statRcvMsgQoS < #MQTT_QOS_2 THEN
                                                           // If QoS is 0 or 1, copy topic directly to output
                                                           #tempReceivedTopicStringMaxLen := MAX_LEN(#receivedTopic);
                                                           IF #statRcvMsgTopicPos <= #tempReceivedTopicStringMaxLen THEN
                                                               #receivedTopic[#statRcvMsgTopicPos] := BYTE_TO_WCHAR(#statRcvBuffer[#tempTrcvBufferPos]);
                                                               #statRcvMsgTopicPos += 1;
                                                           ELSE
                                                               // Max String len reached.
                                                               #statRcvMsgInternalStatus := #MSG_DECODE_STATUS_TOPIC_TOO_LONG;
                                                           END_IF;
                                                       END_IF;

                                                       IF #statRcvMsgQoS = #MQTT_QOS_2 THEN
                                                           // If QoS is 2, copy topic to QoS2 buffer
                                                           IF #statRcvMsgTopicPos <= #MAX_TOPIC_LEN_QOS2 THEN
                                                               #tempReceivedTopic[#statRcvMsgTopicPos] := BYTE_TO_WCHAR(#statRcvBuffer[#tempTrcvBufferPos]);
                                                               #statRcvTopicStorage[#statStoragePos] := #tempReceivedTopic;
                                                               #statRcvMsgTopicPos += 1;
                                                           END_IF;
                                                       END_IF;

                                                       // Decrement topic length and increment buffer position
                                                       #statRcvMsgTopicLen -= 1;
                                                       #tempTrcvBufferPos += 1;

                                                       // Check condition, if topic fully decoded:
                                                       IF #statRcvMsgTopicLen <= 0 THEN
                                                           // Decide what to do next:
                                                           IF #statRcvMsgQoS > #MQTT_QOS_0 THEN
                                                               // NextStep Decode PacketID
                                                               #statRcvMsgDecodeState := #MSG_DECODE_STATE_PACKET_ID_MSB;
                                                           ELSIF #statRcvMsgQoS = #MQTT_QOS_0 AND #statRcvMsgPayloadLen > 0 THEN
                                                               // NextStep Decode Payload
                                                               #statRcvMsgDecodeState := #MSG_DECODE_STATE_PAYLOAD;
                                                           ELSE
                                                               // QoS=0 and no Payload => Done
                                                               // Decoding complete
                                                               #statRcvMsgDecodeState := #MSG_DECODE_STATE_COMPLETED;
                                                           END_IF;
                                                       END_IF;

                                                   #MSG_DECODE_STATE_PACKET_ID_MSB:  // Decode PacketId MSB. Only done if QoS is 1 or 2
                                                       // Copy PacketID
                                                       #statRcvMsgPacketId.%B1 := #statRcvBuffer[#tempTrcvBufferPos]; // MSB
                                                       // Increment buffer position
                                                       #tempTrcvBufferPos += 1; // Increment
                                                       #statRcvMsgDecodeState := #MSG_DECODE_STATE_PACKET_ID_LSB;

                                                   #MSG_DECODE_STATE_PACKET_ID_LSB: // Decode PacketId LSB
                                                       // Copy PacketID
                                                       #statRcvMsgPacketId.%B0 := #statRcvBuffer[#tempTrcvBufferPos]; // LSB
                                                       // If QoS is 2, copy Packet ID to QoS2 buffer
                                                       IF #statRcvMsgQoS = #MQTT_QOS_2 THEN
                                                           #statRcvPacketIdStorage[#statStoragePos] := #statRcvMsgPacketId;
                                                           #tempIntReturn := RD_SYS_T(#statRcvTimestampStorage[#statStoragePos]);
                                                       END_IF;

                                                       // Increment buffer position
                                                       #tempTrcvBufferPos += 1; // Increment

                                                       // Decide what to do next
                                                       IF #statRcvMsgPayloadLen > 0 THEN
                                                           #statRcvMsgDecodeState := #MSG_DECODE_STATE_PAYLOAD;
                                                       ELSE
                                                           // Decoding complete
                                                           #statRcvMsgDecodeState := #MSG_DECODE_STATE_COMPLETED;
                                                       END_IF;

                                                   #MSG_DECODE_STATE_PAYLOAD:
                                                       // Decode Payload
                                                       IF #statRcvMsgQoS < #MQTT_QOS_2 THEN
                                                           // If QoS is 0 or 1, copy payload directly to output
                                                           #tempUpperBoundRcvMsgDataArray := UPPER_BOUND(ARR := #receivedMsgPayload, DIM := #ONE_DIMENSION);
                                                           IF #statRcvMsgPayloadPos <= #tempUpperBoundRcvMsgDataArray THEN
                                                               #receivedMsgPayload[#statRcvMsgPayloadPos] := #statRcvBuffer[#tempTrcvBufferPos];
                                                               #statRcvMsgPayloadPos += 1;
                                                           ELSE
                                                               // Max Payload len reached
                                                               #statRcvMsgInternalStatus := #MSG_DECODE_STATUS_PAYLOAD_TOO_LONG;
                                                           END_IF;
                                                       END_IF;

                                                       IF #statRcvMsgQoS = #MQTT_QOS_2 THEN
                                                           // If QoS is 2, copy payload to QoS2 buffer
                                                           IF #statRcvMsgPayloadPos <= #MAX_BUFFER_LEN_RCV THEN
                                                               #statRcvPayloadStorage[#statStoragePos, #statRcvMsgPayloadPos] := #statRcvBuffer[#tempTrcvBufferPos];
                                                               #statRcvMsgPayloadPos += 1;
                                                           END_IF;
                                                       END_IF;

                                                       // Decrement payload length and increment buffer position
                                                       #statRcvMsgPayloadLen -= 1;
                                                       #tempTrcvBufferPos += 1;

                                                       // Check condition, if payload fully decoded:
                                                       IF #statRcvMsgPayloadLen <= 0 THEN
                                                           // Decoding complete
                                                           #statRcvMsgDecodeState := #MSG_DECODE_STATE_COMPLETED;
                                                       END_IF;

                                                   #MSG_DECODE_STATE_COMPLETED:
                                                       // Write payload length
                                                       IF #statRcvMsgQoS = #MQTT_QOS_2 THEN
                                                           #statRcvMsgPayloadLenStorage[#statStoragePos] := #statDecodedPayloadLenght;
                                                       ELSE
                                                           #tempReceivedMsgDataArrayTotalLen := ABS(UPPER_BOUND(ARR := #receivedMsgPayload, DIM := #ONE_DIMENSION) - LOWER_BOUND(ARR := #receivedMsgPayload, DIM := #ONE_DIMENSION)) + #ARRAY_LEN_OFFSET_PLUS_1;
                                                           IF #statDecodedPayloadLenght > #tempReceivedMsgDataArrayTotalLen THEN
                                                               #statRcvMsgDataLen := DINT_TO_UDINT(#tempReceivedMsgDataArrayTotalLen);
                                                           ELSE
                                                               #statRcvMsgDataLen := #statDecodedPayloadLenght;
                                                           END_IF;
                                                       END_IF;

                                                       // Set internal status if QoS 0 or 1
                                                       IF #statRcvMsgQoS < #MQTT_QOS_2
                                                           AND #statRcvMsgInternalStatus = #MSG_DECODE_STATUS_NO_NEW_MSG
                                                       THEN
                                                           #statRcvMsgInternalStatus := #MSG_DECODE_STATUS_NEW_MSG_OK;
                                                       END_IF;

                                                       // Depending on the QoS of the last received message, send ACK, PUBREC or nothing
                                                       CASE #statRcvMsgQoS OF
                                                           #MQTT_QOS_0:
                                                               #statSendPubRecMsg := FALSE;
                                                               #statSendPubAckMsg := FALSE;
                                                           #MQTT_QOS_1:
                                                               #statSendPubRecMsg := FALSE;
                                                               #statSendPubAckMsg := TRUE;
                                                           #MQTT_QOS_2:
                                                               #statSendPubRecMsg := TRUE;
                                                               #statSendPubAckMsg := FALSE;
                                                       END_CASE;

                                                       // Finish processing
                                                       #statRcvMsgDecodeState := #MSG_DECODE_STATE_NO_PROCESSING;
                                                   ELSE
                                                       // else case
                                                       #statStatus := #ERR_UNDEFINED_STATE;
                                                       #statErrorUserCleared := TRUE;
                                               END_CASE;
                                           END_REGION RECEIVED_PACKET_DECODE

                                       ELSE
                                           // No Header found, SKIP entry of buffer:
                                           #tempTrcvBufferPos += 1;
                                   END_CASE;
                               END_WHILE;

                               REGION POST-PROCESSING OF RECEIVED MESSAGES
                                   // Do post-processing if the processing has finished and there is a message to show
                                   IF #statRcvMsgInternalStatus <> #MSG_DECODE_STATUS_NO_NEW_MSG
                                       AND #statRcvMsgDecodeState = #MSG_DECODE_STATE_NO_PROCESSING
                                   THEN
                                       // Set New message flag
                                       #statRcvMsgStatus := #statRcvMsgInternalStatus;
                                       // Reset internal status
                                       #statRcvMsgInternalStatus := #MSG_DECODE_STATUS_NO_NEW_MSG;
                                   END_IF;
                               END_REGION

                           END_REGION TRCV_NEW_DATA
                       END_IF;

                       // Send an Publish Acknowledge Msg, if necessary
                       REGION SEND_PUBACK_MSG_ON_SUBSCRIPTIONS
                           // Send Acknowledgements to Subscribed messages, if requested (QoS =1)
                           IF #statSendPubAckMsg = TRUE AND // send pub ack Request
                               #statMqttCommandState = #MQTT_COMMAND_STATE_NO_PROCESSING AND // no send job processing
                               #statRcvMsgDecodeState = #MSG_DECODE_STATE_NO_PROCESSING AND // processing of received messages has finished
                               #statTsendcReq = FALSE AND // Not another active send request
                               #tempTsendcBusy = FALSE AND // tsendC is ready
                               #tempTsendcDone = FALSE // tsendC did not finished in this cycle
                           THEN
                               // Set Pos
                               #statSendBufferPos := 0;
                               // Write Msg Type
                               #statSendBuffer[#statSendBufferPos] := #MQTT_MSG_TYPE_PUBACK;
                               #statSendBufferPos += 1;
                               // Write Msg Len
                               #statSendBuffer[#statSendBufferPos] := #REMAINING_LEN_2;
                               #statSendBufferPos += 1;
                               // Write Packet Id - first MSB then LSB
                               #statSendBuffer[#statSendBufferPos] := #statRcvMsgPacketId.%B1;
                               #statSendBufferPos += 1;
                               #statSendBuffer[#statSendBufferPos] := #statRcvMsgPacketId.%B0;
                               #statSendBufferPos += 1;
                               // Set Send Len:
                               #statTsendcLen := #statSendBufferPos;
                               // Send msg
                               #statTsendcReq := TRUE;
                               // Reset ack:
                               #statSendPubAckMsg := FALSE;
                           END_IF;
                       END_REGION SEND_PUBACK_MSG_ON_SUBSCRIPTIONS

                       // Send an Publish Recieved Msg, if necessary
                       REGION SEND_PUBREC_MSG_ON_SUBSCRIPTIONS
                           // Send PUBREC to Subscribed messages, if requested (QoS = 2)
                           IF #statSendPubRecMsg = TRUE AND // send PUBREC
                               #statMqttCommandState = #MQTT_COMMAND_STATE_NO_PROCESSING AND // no send job processing
                               #statRcvMsgDecodeState = #MSG_DECODE_STATE_NO_PROCESSING AND // processing of received messages has finished
                               #statTsendcReq = FALSE AND // Not another active send request
                               #tempTsendcBusy = FALSE AND // tsendC is ready
                               #tempTsendcDone = FALSE // tsendC did not finished in this cycle
                           THEN
                               // Set Pos
                               #statSendBufferPos := 0;
                               // Write Msg Type
                               #statSendBuffer[#statSendBufferPos] := #MQTT_MSG_TYPE_PUBREC;
                               #statSendBufferPos += 1;
                               // Write Msg Len
                               #statSendBuffer[#statSendBufferPos] := #REMAINING_LEN_2;
                               #statSendBufferPos += 1;
                               // Write Packet Id - first MSB then LSB

                               #statSendBuffer[#statSendBufferPos] := #statRcvMsgPacketId.%B1;
                               #statSendBufferPos += 1;
                               #statSendBuffer[#statSendBufferPos] := #statRcvMsgPacketId.%B0;
                               #statSendBufferPos += 1;
                               // Set Send Len:
                               #statTsendcLen := #statSendBufferPos;
                               // Send msg
                               #statTsendcReq := TRUE;
                               // Reset ack:
                               #statSendPubRecMsg := FALSE;
                           END_IF;
                       END_REGION SEND_PUBREC_MSG_ON_SUBSCRIPTIONS

                       // Send an Publish Complete Msg, if necessary
                       REGION SEND_PUBCOMP_MSG_ON_SUBSCRIPTIONS
                           // Send PUBCOM to subscribed messages
                           IF #statSendPubCompMsg = TRUE AND // send pub ack Request
                               #statMqttCommandState = #MQTT_COMMAND_STATE_NO_PROCESSING AND // no send job processing
                               #statTsendcReq = FALSE AND // Not another active send request
                               #tempTsendcBusy = FALSE AND // tsendC is ready
                               #tempTsendcDone = FALSE // tsendC did not finished in this cycle
                           THEN
                               // Set Pos
                               #statSendBufferPos := 0;
                               // Write Msg Type
                               #statSendBuffer[#statSendBufferPos] := #MQTT_MSG_TYPE_PUBCOMP;
                               #statSendBufferPos += 1;
                               // Write Msg Len
                               #statSendBuffer[#statSendBufferPos] := #REMAINING_LEN_2;
                               #statSendBufferPos += 1;
                               // Write Packet Id - first MSB then LSB
                               #statSendBuffer[#statSendBufferPos] := #statRelPacketId.%B1;
                               #statSendBufferPos += 1;
                               #statSendBuffer[#statSendBufferPos] := #statRelPacketId.%B0;
                               #statSendBufferPos += 1;
                               // Set Send Len:
                               #statTsendcLen := #statSendBufferPos;
                               // Send msg
                               #statTsendcReq := TRUE;
                               // Reset PUBCOMP send message:
                               #statSendPubCompMsg := FALSE;
                           END_IF;
                       END_REGION SEND_PUBCOMP_MSG_ON_SUBSCRIPTIONS

                       // MQTT Commands state machine
                       REGION MQTT_STATE_MACHINE
                           CASE #statMqttConnectState OF
                               #MQTT_CONNECT_STATE_NO_PROCESSING:
                                   ;
                               #MQTT_CONNECT_STATE_BUILD_PACKET:
                                   REGION BUILD_CONNECT_PACKET
                                       // Remaining Length is the length of the variable header (10 bytes) plus the length of the Payload. 
                                       // Max Len of Mqtt packets is per Standard 268,435,455 Bytes (ff,ff,ff,7f)
                                       // Calculate Remain Len will be 10 bytes
                                       // plus Len of ClientId   (max 3*16382 WChars= 49.146 Bytes)
                                       // plus Len of User (max 3*16382 WChars= 49.146 Bytes)
                                       // plus Len of PW (max 3*16382 WChars= 49.146 Bytes)
                                       // plus Len of WillTopic (max 3*16382 WChars= 49.146 Bytes)
                                       // plus Len of WillMessage (max 65535 Bytes - as only 2 Bytes Len info is possible)
                                       // = Total 262 119 Bytes


                                       // Must obey, if not currently sending PubAck Msg on a subscription
                                       // Else, try in the next cycle
                                       IF #tempTsendcBusy = FALSE AND // tsendC is ready
                                           #tempTsendcDone = FALSE AND  // tsendC did not finish in this cycle
                                           #statTsendcReq = FALSE THEN // no request from pub ack request

                                           // Only need to encode header once
                                           IF #statPacketHeaderEncodeDone = FALSE THEN
                                               // INIT
                                               #statSendBufferPos := 0;
                                               #statClientIdPos := #FIRST_CHARACTER;
                                               #statClientIdEncodeState := #FIRST_ENCODING;

                                               #statWillTopicEncodeState := #FIRST_ENCODING;
                                               #statWillTopicPos := #FIRST_CHARACTER;

                                               #statWillMessageEncodeState := #FIRST_ENCODING;
                                               #statWillMessagePos := 0; // The Posistion for the WILL Message Array

                                               #statUserNameEncodeState := #FIRST_ENCODING;
                                               #statUserNamePos := #FIRST_CHARACTER;

                                               #statPasswordEncodeState := #FIRST_ENCODING;
                                               #statPasswordPos := #FIRST_CHARACTER;

                                               #statSendPacketTotalRemLen := #CONNECT_HEADER_10BYTE_LEN;
                                               #statClientIdLenUtf8Encoded := 0;
                                               #statWillTopicLenUtf8Encoded := 0;
                                               #statUsernameLenUtf8Encoded := 0;
                                               #statPasswordLenUtf8Encoded := 0;
                                               // End Init

                                               // Encode Client ID Len
                                               // Client ID must always be present
                                               FOR #tempLoopCounter := #FIRST_CHARACTER TO LEN(#clientIdentifier) DO
                                                   "LMQTT_ConvertToUtf8"(character := #clientIdentifier[#tempLoopCounter],
                                                                         convertedUtf8 => #tempConvertedUtf8,
                                                                         bytesUsed => #tempBytesUsedUtf8,
                                                                         error => #tempErrorConvertUtf8,
                                                                         status => #tempStatusConvertUtf8);
                                                   #statClientIdLenUtf8Encoded := #statClientIdLenUtf8Encoded + #tempBytesUsedUtf8;
                                               END_FOR;

                                               #statSendPacketTotalRemLen := #statSendPacketTotalRemLen + #statClientIdLenUtf8Encoded + #TWO_BYTE_LEN_INFO;


                                               IF #username <> #EMPTY_WSTRING THEN
                                                   #tempUserFlag := TRUE;
                                                   FOR #tempLoopCounter := #FIRST_CHARACTER TO LEN(#username) DO
                                                       "LMQTT_ConvertToUtf8"(character := #username[#tempLoopCounter],
                                                                             convertedUtf8 => #tempConvertedUtf8,
                                                                             bytesUsed => #tempBytesUsedUtf8,
                                                                             error => #tempErrorConvertUtf8,
                                                                             status => #tempStatusConvertUtf8);
                                                       #statUsernameLenUtf8Encoded := #statUsernameLenUtf8Encoded + #tempBytesUsedUtf8;
                                                   END_FOR;
                                                   #statSendPacketTotalRemLen := #statSendPacketTotalRemLen + #statUsernameLenUtf8Encoded + #TWO_BYTE_LEN_INFO;
                                               ELSE
                                                   #statUserNameEncodeState := #NOT_USED_NO_ENCODING;
                                                   #tempUserFlag := FALSE;
                                               END_IF;

                                               IF #password <> #EMPTY_WSTRING AND #username <> #EMPTY_WSTRING THEN
                                                   #tempPasswordFlag := TRUE;
                                                   FOR #tempLoopCounter := #FIRST_CHARACTER TO LEN(#password) DO
                                                       "LMQTT_ConvertToUtf8"(character := #password[#tempLoopCounter],
                                                                             convertedUtf8 => #tempConvertedUtf8,
                                                                             bytesUsed => #tempBytesUsedUtf8,
                                                                             error => #tempErrorConvertUtf8,
                                                                             status => #tempStatusConvertUtf8);
                                                       #statPasswordLenUtf8Encoded := #statPasswordLenUtf8Encoded + #tempBytesUsedUtf8;
                                                   END_FOR;
                                                   #statSendPacketTotalRemLen := #statSendPacketTotalRemLen + #statPasswordLenUtf8Encoded + #TWO_BYTE_LEN_INFO;
                                               ELSE
                                                   #statPasswordEncodeState := #NOT_USED_NO_ENCODING;
                                                   #tempPasswordFlag := FALSE;
                                               END_IF;


                                               IF #willtopic <> #EMPTY_WSTRING THEN
                                                   #tempWillFlag := TRUE;
                                                   CASE #statWillQos OF
                                                       #MQTT_QOS_0:  // Statement section case 1
                                                           #tempWillQoS1 := FALSE;
                                                           #tempWillQoS2 := FALSE;
                                                       #MQTT_QOS_1:  // Statement section case 2 to 4
                                                           #tempWillQoS1 := TRUE;
                                                           #tempWillQoS2 := FALSE;
                                                       #MQTT_QOS_2:
                                                           #tempWillQoS1 := FALSE;
                                                           #tempWillQoS2 := True;
                                                       ELSE  // Statement section ELSE
                                                           ;
                                                   END_CASE;
                                                   FOR #tempLoopCounter := #FIRST_CHARACTER TO LEN(#willtopic) DO
                                                       // Statement section FOR
                                                       "LMQTT_ConvertToUtf8"(character := #willtopic[#tempLoopCounter],
                                                                             convertedUtf8 => #tempConvertedUtf8,
                                                                             bytesUsed => #tempBytesUsedUtf8,
                                                                             error => #tempErrorConvertUtf8,
                                                                             status => #tempStatusConvertUtf8);
                                                       #statWillTopicLenUtf8Encoded := #statWillTopicLenUtf8Encoded + #tempBytesUsedUtf8;
                                                   END_FOR;
                                                   // Add WillTopic Len and Will Message Len (and len info twice)
                                                   #statSendPacketTotalRemLen := #statSendPacketTotalRemLen + #statWillTopicLenUtf8Encoded + #statWillMessageCnt + (2 * #TWO_BYTE_LEN_INFO);
                                               ELSE
                                                   #statWillTopicEncodeState := #NOT_USED_NO_ENCODING;
                                                   #statWillMessageEncodeState := #NOT_USED_NO_ENCODING;
                                                   #tempWillFlag := FALSE;
                                                   #statWillRetain := FALSE;
                                                   #tempWillQoS1 := FALSE;
                                                   #tempWillQoS2 := FALSE;
                                               END_IF;

                                               // Build Connect Telegram
                                               // Fixed Header - Write Packet Type
                                               #statSendBuffer[#statSendBufferPos] := #MQTT_MSG_TYPE_CONNECT; // 1 Byte
                                               #statSendBufferPos += 1; // increment

                                               // Write Remaining Packet Len info 
                                               WHILE (#statSendPacketTotalRemLen > #DEFAULT_VALUE_ZERO)
                                               DO// See MQTT Spec for explanation of this calculation
                                                   #statEncodedRemPacketLenAsByte := UDINT_TO_BYTE(#statSendPacketTotalRemLen MOD #SEND_LEN_MULTIPLIER_UDINT_128);
                                                   #statSendPacketTotalRemLen := #statSendPacketTotalRemLen / #SEND_LEN_MULTIPLIER_UDINT_128;
                                                   // if there are more data to encode, set the top bit of this byte
                                                   IF #statSendPacketTotalRemLen > #DEFAULT_VALUE_ZERO THEN
                                                       // Do this and continue while loop
                                                       #statEncodedRemPacketLenAsByte := #statEncodedRemPacketLenAsByte OR UDINT_TO_BYTE(#SEND_LEN_MULTIPLIER_UDINT_128);
                                                       #statSendBuffer[#statSendBufferPos] := #statEncodedRemPacketLenAsByte;
                                                       #statSendBufferPos += 1;
                                                   ELSE
                                                       // Do this and leave while loop
                                                       #statSendBuffer[#statSendBufferPos] := #statEncodedRemPacketLenAsByte;
                                                       #statSendBufferPos += 1;
                                                   END_IF;
                                               END_WHILE;

                                               // Build Connect Telegram
                                               // Write Protocol name
                                               #statSendBuffer[#statSendBufferPos] := #CONN_PROTOCOL_NAME_0;
                                               #statSendBufferPos += 1;
                                               #statSendBuffer[#statSendBufferPos] := #CONN_PROTOCOL_NAME_4;
                                               #statSendBufferPos += 1;
                                               #statSendBuffer[#statSendBufferPos] := CHAR_TO_BYTE('M');
                                               #statSendBufferPos += 1;
                                               #statSendBuffer[#statSendBufferPos] := CHAR_TO_BYTE('Q');
                                               #statSendBufferPos += 1;
                                               #statSendBuffer[#statSendBufferPos] := CHAR_TO_BYTE('T');
                                               #statSendBufferPos += 1;
                                               #statSendBuffer[#statSendBufferPos] := CHAR_TO_BYTE('T');
                                               #statSendBufferPos += 1;
                                               // Write Protocol Level
                                               #statSendBuffer[#statSendBufferPos] := #CONN_PROTOCOL_MQTT_VERSION_3_1_1;
                                               #statSendBufferPos += 1;
                                               // Write Connect Flags
                                               #statSendBuffer[#statSendBufferPos].%X0 := false;
                                               #statSendBuffer[#statSendBufferPos].%X1 := #cleanSession;
                                               #statSendBuffer[#statSendBufferPos].%X2 := #tempWillFlag;
                                               #statSendBuffer[#statSendBufferPos].%X3 := #tempWillQoS1;
                                               #statSendBuffer[#statSendBufferPos].%X4 := #tempWillQoS2;
                                               #statSendBuffer[#statSendBufferPos].%X5 := #statWillRetain;
                                               #statSendBuffer[#statSendBufferPos].%X6 := #tempPasswordFlag;
                                               #statSendBuffer[#statSendBufferPos].%X7 := #tempUserFlag;
                                               #statSendBufferPos += 1;
                                               // Write Keep Alive in sec
                                               #tempWordForSliceAddress := UINT_TO_WORD(#connParam.keepAlive);
                                               #statSendBuffer[#statSendBufferPos] := #tempWordForSliceAddress.%B1;
                                               #statSendBufferPos += 1;
                                               #statSendBuffer[#statSendBufferPos] := #tempWordForSliceAddress.%B0;
                                               #statSendBufferPos += 1;

                                               // Set To Complete this, can skip in further progess
                                               #statPacketHeaderEncodeDone := TRUE;
                                           END_IF;

                                           // Payload
                                           // These fields, if present, MUST appear in the order:
                                           // Client Identifier, Will topic, Will message, User Name, password


                                           // ClientIdentifier
                                           IF #statSendBufferPos <= #MAX_BUFFER_LEN_SEND - #TWO_BYTE_LEN_INFO THEN
                                               CASE #statClientIdEncodeState OF
                                                   #FIRST_ENCODING:  // Statement section case 1
                                                       // ADD len info into packet

                                                       #tempWordForSliceAddress := UINT_TO_WORD(#statClientIdLenUtf8Encoded);
                                                       #statSendBuffer[#statSendBufferPos] := #tempWordForSliceAddress.%B1; // MSB
                                                       #statSendBufferPos += 1;
                                                       #statSendBuffer[#statSendBufferPos] := #tempWordForSliceAddress.%B0; // LSB
                                                       #statSendBufferPos += 1;

                                                       FOR #tempLoopCounter := #statClientIdPos TO LEN(#clientIdentifier) DO
                                                           "LMQTT_ConvertToUtf8"(character := #clientIdentifier[#tempLoopCounter],
                                                                                 convertedUtf8 => #tempConvertedUtf8,
                                                                                 bytesUsed => #tempBytesUsedUtf8,
                                                                                 error => #tempErrorConvertUtf8,
                                                                                 status => #tempStatusConvertUtf8);

                                                           IF #statSendBufferPos + #tempBytesUsedUtf8 <= #MAX_BUFFER_LEN_SEND THEN
                                                               #statClientIdPos += 1;
                                                               CASE #tempBytesUsedUtf8 OF
                                                                   #UTF_1_BYTE_USED:  // Statement section case 1
                                                                       #statSendBuffer[#statSendBufferPos] := #tempConvertedUtf8.%B0;
                                                                       #statSendBufferPos += 1;
                                                                   #UTF_2_BYTE_USED:
                                                                       #statSendBuffer[#statSendBufferPos] := #tempConvertedUtf8.%B0;
                                                                       #statSendBufferPos += 1;
                                                                       #statSendBuffer[#statSendBufferPos] := #tempConvertedUtf8.%B1;
                                                                       #statSendBufferPos += 1;
                                                                   #UTF_3_BYTE_USED:  // Statement section case 2 to 4
                                                                       #statSendBuffer[#statSendBufferPos] := #tempConvertedUtf8.%B0;
                                                                       #statSendBufferPos += 1;
                                                                       #statSendBuffer[#statSendBufferPos] := #tempConvertedUtf8.%B1;
                                                                       #statSendBufferPos += 1;
                                                                       #statSendBuffer[#statSendBufferPos] := #tempConvertedUtf8.%B2;
                                                                       #statSendBufferPos += 1;
                                                                   ELSE  // Statement section ELSE
                                                                       ;
                                                               END_CASE;
                                                           ELSE
                                                               // When buffer full
                                                               #statClientIdEncodeState := #SUBSEQUENT_ENCODING;
                                                               EXIT;
                                                           END_IF;
                                                       END_FOR;
                                                       IF #statClientIdPos >= LEN(#clientIdentifier) THEN
                                                           #statClientIdEncodeState := #ENCODE_DONE;
                                                       END_IF;


